(* IEC 61131-3 sources: kns-port-domestic/upstream/kns-pump-station/src/POUs/Model/F_FaultInjEqual, 2 files *)

(* ---- F_FaultInjEqual.decl.st ---- *)
// Назначение: сравнение двух наборов инъекций ST_FaultInjection поле за полем (структуры в CODESYS
//             оператором «=» не сравниваются; поля REAL — по битам, чтобы NaN был равен NaN).
//             FB_PlantModel по нему считает изменения инъекций
//             (stSimSts.udiFaultSeq → событие журнала 101021). Новое поле ST_FaultInjection добавляется
//             и сюда — тест FaultSeqCountsChanges меняет каждое поле.
// Автор:      kr0nsch
// Версия:     0.1.1
// Документ:   docs/DESIGN.md, разделы 3.3, 11.1
FUNCTION F_FaultInjEqual : BOOL
VAR_IN_OUT CONSTANT
    stA : ST_FaultInjection;
    stB : ST_FaultInjection;
END_VAR
VAR
    uiI : UINT;             // индекс насоса или датчика
    uBitsA : PL.U_RealBits; // поле REAL набора A как биты (сравнение NaN)
    uBitsB : PL.U_RealBits;
END_VAR

(* ---- F_FaultInjEqual.impl.st ---- *)
F_FaultInjEqual := FALSE;
FOR uiI := 1 TO GVL_Const.STN_PUMP_COUNT DO
    IF stA.axVfdFault[uiI] <> stB.axVfdFault[uiI] OR stA.axNoFeedback[uiI] <> stB.axNoFeedback[uiI]
       OR stA.axFeedbackStuck[uiI] <> stB.axFeedbackStuck[uiI] OR stA.axAirLock[uiI] <> stB.axAirLock[uiI]
       OR stA.axClog[uiI] <> stB.axClog[uiI] OR stA.axOverheat[uiI] <> stB.axOverheat[uiI]
       OR stA.axLeak[uiI] <> stB.axLeak[uiI] OR stA.axVfdCommLoss[uiI] <> stB.axVfdCommLoss[uiI]
       OR stA.axLocal[uiI] <> stB.axLocal[uiI] OR stA.axLocalRun[uiI] <> stB.axLocalRun[uiI] THEN
        RETURN;
    END_IF
END_FOR
// поля REAL — по битам (U_RealBits): NaN = NaN, иначе записанный NaN давал бы «изменение» в каждом вызове
FOR uiI := 1 TO GVL_Const.SIM_AI_COUNT DO
    uBitsA.rValue := stA.arAiForced_mA[uiI];
    uBitsB.rValue := stB.arAiForced_mA[uiI];
    IF stA.aeAiFault[uiI] <> stB.aeAiFault[uiI] OR uBitsA.dwValue <> uBitsB.dwValue THEN
        RETURN;
    END_IF
END_FOR
IF stA.eLs102Stuck <> stB.eLs102Stuck OR stA.eLs103Stuck <> stB.eLs103Stuck OR stA.xPowerLoss <> stB.xPowerLoss
   OR stA.xUpsFault <> stB.xUpsFault OR stA.xTempCommLoss <> stB.xTempCommLoss OR stA.xFanFault <> stB.xFanFault
   OR stA.xFanNoFeedback <> stB.xFanNoFeedback OR stA.xValveChamberFlood <> stB.xValveChamberFlood
   OR stA.xFire <> stB.xFire THEN
    RETURN;
END_IF
uBitsA.rValue := stA.rH2S_mgm3;
uBitsB.rValue := stB.rH2S_mgm3;
IF uBitsA.dwValue <> uBitsB.dwValue THEN
    RETURN;
END_IF
uBitsA.rValue := stA.rCh4_pctLel;
uBitsB.rValue := stB.rCh4_pctLel;
IF uBitsA.dwValue <> uBitsB.dwValue THEN
    RETURN;
END_IF
F_FaultInjEqual := TRUE;
